Fanuc KAREL source: MP0169.KL

PROGRAM MP0169
%STACKSIZE=65535
%PRIORITY=65535
%NOLOCKGROUP
ROUTINE FINT(P1 : INTEGER) : INTEGER FROM MP0169
ROUTINE FREAL(P1 : REAL) : REAL FROM MP0169
ROUTINE RTEST(P1 : INTEGER; P2 : REAL) FROM MP0169
ROUTINE FINT
BEGIN
RETURN((P1 + 1))
END FINT
ROUTINE FREAL
BEGIN
RETURN((P1 + 1.0))
END FREAL
ROUTINE RTEST
VAR
U2C_1 : INTEGER
U2C_2 : INTEGER
U2C_3 : INTEGER
U2C_4 : INTEGER
U2C_5 : INTEGER
U2C_6 : INTEGER
S1 : INTEGER
U2C_8 : REAL
BEGIN
U2C_1=7
U2C_2=3
U2C_3=2
U2C_4=1075838976
U2C_5=1083179008
U2C_6=1069547520
-- UNRESOLVED_PC line 28 opcodes [27 27 21 21 21 6B 69 76 23] marker_code=162
END RTEST
BEGIN
RTEST(7,2.5)
END MP0169
